{region 'Documentation'}
(*!
<summary>Checks inequality with the forbidden UDINT value.</summary>
*)
{endregion}
FUNCTION_BLOCK AssertNotEqual_UDInt EXTENDS AssertionBase
VAR_INPUT
    IN : UDINT; //! Actual value checked or observed by this Assertion.
    Expected : UDINT; //! Value that must differ from IN under this Assertion's comparison rules.
END_VAR

SUPER^();

{region 'Documentation'}
(*!
<summary>Check inequality with the forbidden UDINT value.</summary>
*)
{endregion}
METHOD PROTECTED Assert
VAR
    Message : STRING(GVL_Constants.MessageLength);
    ExpectedText : STRING(GVL_Constants.AssertionValueLength);
    ActualText : STRING(GVL_Constants.AssertionValueLength);
END_VAR
IF NOT EvaluationActive THEN
    RETURN;
END_IF;

IF Result = E_Result.Error THEN
    RETURN;
END_IF;

IF Result = E_Result.Failed THEN
    RETURN;
END_IF;

IF IN = Expected THEN
    ExpectedText := UDINT_TO_STRING(Expected);
    ActualText := UDINT_TO_STRING(IN);
    Message := CONCAT('Assertion failed: values are equal but should differ. NotExpected = ',
        ExpectedText);
    Message := CONCAT(Message, ', Actual = ');
    Message := CONCAT(Message, ActualText);
    Message := CONCAT(Message, '.');
    Fail(Message := Message);
    RETURN;
END_IF;

Pass();
END_METHOD

END_FUNCTION_BLOCK

(* stored: Version 1.1.0.1
   POU AssertNotEqual_UDInt: Id {63c66cfa-59ac-4182-b2ab-559c7b3fbbc2}, SpecialFunc None
   Folder Internal: Id {6711f952-87c0-4b13-9d2f-b610188ec8a0}
   Method Assert: Id {98944a14-deb1-45c1-b066-a31f9ba1de1d} *)
